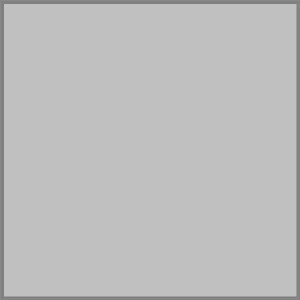
VISUALIZATION viz_HMI_LockIndex  // 300x300
    Rectangle (0,0 300x300), invisible if: not prg_HMI_OperationLock.b_LockIndex
END_VISUALIZATION

(* stored: Version 1.1.0.1, ProductVersion 3.1.4024.13
   Visu viz_HMI_LockIndex: Id {282ec89c-e3f2-491b-b960-931638ae7c1b} *)
